(* LS Electric XG5000 project: TX00N *)
(* PLC LSPLC *)

PROGRAM NewProgram (* task: 스캔 프로그램 *)
VAR
    Count : LINT; (* Source preservation check *)
END_VAR
Count := Count + 1;
END_PROGRAM

PROGRAM AddedST (* task: 스캔 프로그램 *)
VAR
    Count : LINT; (* Source preservation check *)
END_VAR
Count := Count + 1;
END_PROGRAM